// TIA Portal V21 export
// export: Created 2026-11-10T23:32:32.7566402Z, ExportSetting WithDefaults, DisplayName Totally Integrated Automation Portal, DisplayVersion V21 Update 3, DisplayName STEP 7 Professional, DisplayVersion V21 Update 3, DisplayName STEP 7 Safety, DisplayVersion V21, DisplayName Tech WebApplication, DisplayVersion V21, DisplayName WinCC Basic/Comfort/Advanced, DisplayVersion V21 Update 3, DisplayName WinCC Unified, DisplayVersion V21 Update 3
DATA_BLOCK "mTO_Kinematics"   // DB6, Motion_DB
// stored: AutoNumber true, DBAccessibleFromOPCUA true, DBAccessibleFromWebserver true, InstanceOfName TO_Kinematics, OfSystemLibElement TO_Kinematics, OfSystemLibVersion 8.0
TO_Kinematics   // technology object, version 8.0
// stored: KinematicsAxis Ref mTO_PositioningAxis, Type TO_PositioningAxis, Index 1
// stored: KinematicsAxis Ref mTO_SynchronousAxis, Type TO_SynchronousAxis, Index 2
   // // inherited from TO_Object
   // VAR
   //    Tcp { ExternalWritable := 'False'; S7_SetPoint := 'True'} : TO_Struct_Kinematics_StatusKinematicsFrameTcp;
   //    Kinematics { S7_SetPoint := 'True'} : TO_Struct_Kinematics_Kinematics;
   //    KcsFrame { S7_SetPoint := 'True'} : TO_Struct_Kinematics_Frame;
   //    OcsFrame { S7_SetPoint := 'True'} : Array[1..3] of TO_Struct_Kinematics_Frame;
   //    Tool { S7_SetPoint := 'True'} : Array[1..3] of TO_Struct_Kinematics_Tool;
   //    DynamicDefaults { S7_SetPoint := 'True'} : TO_Struct_Kinematics_DynamicDefaults;
   //    DynamicLimits { S7_SetPoint := 'True'} : TO_Struct_Kinematics_DynamicLimits;
   //    Joint { S7_SetPoint := 'True'} : TO_Struct_Kinematics_Joint;
   //    AxisCoupling { S7_SetPoint := 'True'} : TO_Struct_Kinematics_AxisCoupling;
   //    MotionQueue { ExternalWritable := 'False'; S7_SetPoint := 'True'} : TO_Struct_Kinematics_MotionQueue;
   //    Transition { S7_SetPoint := 'True'} : TO_Struct_Kinematics_Transition;
   //    Override { S7_SetPoint := 'True'} : TO_Struct_Kinematics_Override;
   //    Conveyor { S7_SetPoint := 'True'} : TO_Struct_Kinematics_Conveyor;
   //    WorkspaceZone { S7_SetPoint := 'True'} : Array[1..10] of TO_Struct_Kinematics_WorkSpaceZone;
   //    KinematicsZone { S7_SetPoint := 'True'} : Array[2..10] of TO_Struct_Kinematics_KinematicsZone;
   //    StatusPath { ExternalWritable := 'False'; S7_SetPoint := 'True'} : TO_Struct_Kinematics_StatusPath;
   //    TcpInWcs { ExternalWritable := 'False'; S7_SetPoint := 'True'} : TO_Struct_Kinematics_StatusKinematicsFrameWithDynamics;
   //    TcpInOcs { ExternalWritable := 'False'; S7_SetPoint := 'True'} : Array[1..3] of TO_Struct_Kinematics_StatusKinematicsFrameWithDynamicsOcs;
   //    StatusOcsFrame { ExternalWritable := 'False'; S7_SetPoint := 'True'} : Array[1..3] of TO_Struct_Kinematics_StatusFrame;
   //    StatusKinematics { ExternalWritable := 'False'; S7_SetPoint := 'True'} : TO_Struct_Kinematics_StatusKinematics;
   //    AxesData { ExternalWritable := 'False'; S7_SetPoint := 'True'} : TO_Struct_Kinematics_AxesData;
   //    JointData { ExternalWritable := 'False'; S7_SetPoint := 'True'} : TO_Struct_Kinematics_StatusJointData;
   //    FlangeInKcs { ExternalWritable := 'False'; S7_SetPoint := 'True'} : TO_Struct_Kinematics_StatusFlangeInKcs;
   //    StatusTool { ExternalWritable := 'False'; S7_SetPoint := 'True'} : TO_Struct_Kinematics_StatusTool;
   //    StatusConveyor { ExternalWritable := 'False'; S7_SetPoint := 'True'} : Array[1..3] of TO_Struct_Kinematics_StatusConveyor;
   //    StatusWorkspaceZone { ExternalWritable := 'False'; S7_SetPoint := 'True'} : Array[1..10] of TO_Struct_Kinematics_StatusWorkSpaceZone;
   //    StatusKinematicsZone { ExternalWritable := 'False'; S7_SetPoint := 'True'} : Array[2..10] of TO_Struct_Kinematics_StatusKinematicsZone;
   //    StatusZoneMonitoring { ExternalWritable := 'False'; S7_SetPoint := 'True'} : TO_Struct_Kinematics_StatusZoneMonitoring;
   //    StatusMotionQueue { ExternalWritable := 'False'; S7_SetPoint := 'True'} : TO_Struct_Kinematics_StatusMotionQueue;
   //    KinematicsAxis { ExternalWritable := 'False'; S7_SetPoint := 'True'} : TO_Struct_Kinematics_KinematicsAxis;
   //    Units { ExternalWritable := 'False'; S7_SetPoint := 'True'} : TO_Struct_Kinematics_Units;
   //    StatusInterpreterMotion { ExternalWritable := 'False'; S7_SetPoint := 'True'} : TO_Struct_Kinematics_StatusInterpreterMotion;
   //    StatusWord { ExternalWritable := 'False'} : DWord;
   //    ErrorWord { ExternalWritable := 'False'} : DWord;
   //    ErrorDetail { ExternalWritable := 'False'; S7_SetPoint := 'True'} : TO_Struct_ErrorDetail;
   //    WarningWord { ExternalWritable := 'False'} : DWord;
   //    ControlPanel { S7_SetPoint := 'True'} : TO_Struct_Kinematics_ControlPanel;
   //    InternalToTrace { S7_SetPoint := 'True'} : Array[1..4] of TO_Struct_Internal;
   // END_VAR
BEGIN
END_DATA_BLOCK
